(* IEC 61131-3 sources: rusty/tests/lit/ir_tests, 10 files *)

(* ---- adr_ptr_arith.st ---- *)
// RUN: %COMPILE_IR %s | %CHECK_IR %s
//
// Structural pin for the #1749 fix: `ADR(x) + N` must lower to
// `ptrtoint` + `add` (byte-stride integer arithmetic), not panic. ADR is
// declared `: LWORD` so the binary `+` flows through the integer path; the
// codegen entry now routes pointer operands through
// `convert_to_int_value_if_pointer` (matching the existing comparison-op
// path) instead of an unconditional `into_int_value()` that crashed inkwell.

FUNCTION main
VAR
    arr : ARRAY[0..3] OF BYTE;
    pt  : REF_TO BYTE;
END_VAR

pt := ADR(arr) + 2;
pt^ := BYTE#16#FF;
END_FUNCTION

// CHECK: ptrtoint ptr %{{.*}} to i64
// CHECK-NEXT: add i64 %{{.*}}, 2
// CHECK-NEXT: inttoptr i64 %{{.*}} to ptr

(* ---- var_input_aggregate_pass_by_ref.st ---- *)
// RUN: %COMPILE_IR %s | %CHECK_IR %s

// Aggregate VAR_INPUT arguments must be passed by pointer; emitting
// `bitcast ptr -> [N x T]` is invalid IR. See #1718.

FUNCTION foo
   VAR_INPUT
       arr : ARRAY[1..3] OF DINT;
   END_VAR
END_FUNCTION

FUNCTION main
   foo([1, 2, 3]);
END_FUNCTION

// CHECK-LABEL: define {{.*}}@main
// CHECK:       %{{[a-zA-Z0-9_.]+}} = alloca [3 x i32]
// CHECK:       store [3 x i32]
// CHECK:       call {{.*}}@foo(ptr {{.*}})
// CHECK-NOT:   bitcast ptr {{.*}} to [

(* ---- variadic_null_terminator.st ---- *)
// RUN: %COMPILE_IR %s | %CHECK_IR %s
//
// Calls to untyped C-style variadics (`args : ...`) carry an implicit null pointer as their
// last argument. The callee has no way of its own to know how many arguments it received, so
// APIs that walk the list until a terminator read past the arguments without it. Format- and
// count-directed callees read only the arguments they expect and never see the terminator.
//
// Typed variadics keep their argument list unchanged: a `{sized} T...` passes (count, array)
// and a typed unsized `T...` has a concrete callee signature, so a terminator would corrupt
// the contract in both cases.

{external}
FUNCTION untyped : DINT
VAR_INPUT
    fmt : STRING;
    args : ...;
END_VAR
END_FUNCTION

{external}
FUNCTION typed : DINT
VAR_INPUT
    count : DINT;
    args : DINT...;
END_VAR
END_FUNCTION

{external}
FUNCTION sized : DINT
VAR_INPUT
    args : {sized} DINT...;
END_VAR
END_FUNCTION

FUNCTION main : DINT
VAR
    text : STRING := 'text';
END_VAR
    // A call without any variadic argument is still terminated. This is the case in which a
    // terminator-based callee reads past the argument list without the terminator.
    untyped(text);
    // CHECK: call i32 (ptr, ...) @untyped(ptr {{.*}}, ptr null)

    untyped(text, DINT#1, DINT#2);
    // CHECK: call i32 (ptr, ...) @untyped(ptr {{.*}}, i32 1, i32 2, ptr null)

    // The `, !dbg` suffix pins the end of the argument list, so an added terminator fails here.
    typed(DINT#2, DINT#1, DINT#2);
    // CHECK: call i32 (i32, ...) @typed(i32 2, i32 1, i32 2), !dbg

    sized(DINT#1, DINT#2, DINT#3);
    // CHECK: call i32 @sized(i32 3, ptr {{.*}}), !dbg
END_FUNCTION

(* ---- action_call_stores_var_in_out_address.st ---- *)
// RUN: %COMPILE_IR %s | %CHECK_IR %s
//
// Pin the IR shape that the #1576 fix (commit 2b3388f) put in place: when
// calling an action that inherits a `VAR_IN_OUT` from its parent FB, the
// caller must (a) GEP to the FB's in-out slot and (b) store the local's
// address there before invoking the action. Skipping either step leaves the
// pointer NULL and the action segfaults at runtime — runtime coverage lives
// in `tests/lit/single/actions/action_call_with_var_in_out.st`; this test
// is the structural guardrail.

PROGRAM mainProg
VAR
    fb : fb_t;
    localBool : BOOL;
END_VAR
    fb.foo(myInOut := localBool);
END_PROGRAM

FUNCTION_BLOCK fb_t
VAR_IN_OUT
    myInOut : BOOL;
END_VAR
END_FUNCTION_BLOCK

ACTIONS
    ACTION foo
        myInOut := myInOut;
    END_ACTION
END_ACTIONS

// CHECK-LABEL: define void @mainProg(
// CHECK: %fb = getelementptr inbounds nuw %mainProg, {{.*}}, i32 0, i32 0
// CHECK: %localBool = getelementptr inbounds nuw %mainProg, {{.*}}, i32 0, i32 1
// CHECK: getelementptr inbounds %fb_t, ptr %fb, i32 0, i32 1
// CHECK-NEXT: store ptr %localBool, ptr {{%[0-9]+}}, align 8
// CHECK-NEXT: call void @fb_t__foo(ptr %fb)

(* ---- external_fb_array_const_init.st ---- *)
// RUN: %COMPILE_IR --generate-external-constructors %s | %CHECK_IR %s
//
// When an {external} function block has an array with a constant initializer,
// compiling with --generate-external-constructors should:
//   1. Produce a .const_init global for the array
//   2. Define (not declare) the ctor
//   3. Use memcpy from the .const_init in the ctor body

{external}
FUNCTION_BLOCK myFb
VAR
    arr : ARRAY[0..4] OF DINT := [1, 2, 3, 4, 5];
END_VAR
END_FUNCTION_BLOCK

PROGRAM Main
VAR
    fb : myFb;
END_VAR
END_PROGRAM

// The const_init global should exist for the array
// CHECK: @.const_init = private unnamed_addr constant [5 x i32] [i32 1, i32 2, i32 3, i32 4, i32 5]

// The ctor for myFb should be defined (has body), not just declared
// CHECK: define void @myFb__ctor(ptr %0)

// The ctor should use memcpy from the const_init
// CHECK: call void @llvm.memcpy{{.*}}@.const_init

(* ---- external_fb_array_no_init_globals.st ---- *)
// RUN: %COMPILE_IR %s | %CHECK_IR %s
//
// When an {external} function block has an array with a constant initializer,
// compiling WITHOUT --generate-external-constructors should:
//   1. NOT produce any .const_init or __init globals for the external FB
//   2. Declare (not define) the ctor

{external}
FUNCTION_BLOCK myFb
VAR
    arr : ARRAY[0..4] OF DINT := [1, 2, 3, 4, 5];
END_VAR
END_FUNCTION_BLOCK

PROGRAM Main
VAR
    fb : myFb;
END_VAR
END_PROGRAM

// No .const_init or __myFb.arr__init globals should be present.
// CHECK-NOT directives must come before CHECK to scan from start of input.
// CHECK-NOT: @.const_init
// CHECK-NOT: @__myFb.arr__init

// The ctor for myFb should be declared (external), not defined
// CHECK: declare void @myFb__ctor(ptr)

(* ---- fb_call_no_int_extension_attrs.st ---- *)
// REQUIRES: host-x86_64
// RUN: %COMPILE_IR %s | %CHECK_IR %s
//
// Direct FUNCTION_BLOCK invocations (e.g. `myFbInstance(in_val := …)`) lower to
// a gep+store of each argument into the instance struct followed by a call to
// the FB body that takes only the instance pointer — there are no scalar
// arguments in the LLVM call signature, so no `signext`/`zeroext` attribute is
// applicable. Regression for #1146 review feedback: confirms the call-side
// integer-extension pass leaves direct FB calls alone.
//
// Gated to host-x86_64 to mirror sub32_int_ffi_extension.st: `signext`/`zeroext`
// are only emitted on x86 family and Apple/Darwin targets. The point of this
// test is the *absence* of those tokens, but on AAPCS targets they would be
// absent for a different reason (target gate), which would make the test
// trivially green and hide a future regression on x86.

FUNCTION_BLOCK myFb
VAR_INPUT
    in_val : SINT;
END_VAR
END_FUNCTION_BLOCK

PROGRAM main
VAR
    instance : myFb;
END_VAR
    instance(in_val := SINT#-1);
END_PROGRAM

// The body call passes only the instance struct pointer (LLVM 21 opaque
// `ptr`) — no `signext`/`zeroext` token should appear on the call line.
// CHECK: call void @myFb(ptr {{.*}})
// CHECK-NOT: call void @myFb({{.*}}signext{{.*}})
// CHECK-NOT: call void @myFb({{.*}}zeroext{{.*}})

(* ---- included_struct_ctor.st ---- *)
// RUN: %COMPILE_IR -i %p/include/included_types.st %s | %CHECK_IR %s

PROGRAM Main
VAR
    s : IncludedStruct;
END_VAR
END_PROGRAM

// The declaration may precede or follow Main__ctor depending on the unit order
// CHECK-NOT: define{{.*}}@IncludedStruct__ctor
// CHECK-DAG: define void @Main__ctor(ptr %0) {
// CHECK-DAG: call void @IncludedStruct__ctor(ptr %s)
// CHECK-DAG: declare void @IncludedStruct__ctor(ptr)
// CHECK-NOT: define{{.*}}@IncludedStruct__ctor

(* ---- nested_array_const_expression_init.st ---- *)
// RUN: %COMPILE_IR %s | %CHECK_IR %s
//
// Structural pin for the PRG-4521 fix: constant expressions inside nested
// array initializers are const-folded, so the initializer lowers to a folded
// constant global copied via memcpy. Previously the raw expression tree
// reached codegen's literal generator and failed with "Cannot generate
// Literal for BinaryExpression". Runtime coverage lives in
// tests/lit/single/init/array_const_expression_init.st.

PROGRAM mainProg
VAR
    mArr : ARRAY[0..1] OF ARRAY[0..1] OF UDINT := [[UDINT#0 + UDINT#1, UDINT#0], [UDINT#0, UDINT#2 - UDINT#1]];
END_VAR
    ;
END_PROGRAM

// The type's __init global is fully folded to [1, 0], [0, 1].
// CHECK: @__mainProg.mArr__init = unnamed_addr constant [2 x [2 x i32]] {{\[}}[2 x i32] [i32 1, i32 0], [2 x i32] [i32 0, i32 1]]

// The ctor assignment is folded as well and copied via memcpy.
// CHECK: @.const_init = private unnamed_addr constant [2 x [2 x i32]] {{\[}}[2 x i32] [i32 1, i32 0], [2 x i32] [i32 0, i32 1]]
// CHECK: define void @mainProg__ctor(ptr %0)
// CHECK: call void @llvm.memcpy{{.*}}@.const_init

(* ---- sub32_int_ffi_extension.st ---- *)
// REQUIRES: host-x86_64
// RUN: %COMPILE_IR %s | %CHECK_IR %s
//
// Regression for #1146. Verify call sites and declarations of functions taking sub-32-bit
// integer parameters carry the correct LLVM `signext`/`zeroext` parameter attributes.
// Without these, optimized release builds of FFI'd callees (e.g. the Rust stdlib) read
// garbage upper register bits instead of the intended signed value — see also
// `cargo test --release -p iec61131std mul_ltime_signed`.
//
// Gated to host-x86_64 because the codegen emission is target-aware: x86 family and
// Apple/Darwin emit the attributes; plain AAPCS (aarch64-unknown-linux-gnu) does not
// and the FILECHECK lines below would not match. The runtime regression coverage for
// the AAPCS path lives under tests/lit/single/stdlib_overflow/sub32_ffi_return_*.st.

{external}
FUNCTION extFunc : LINT
VAR_INPUT
    in1 : SINT;
    in2 : USINT;
    in3 : INT;
    in4 : UINT;
    in5 : BOOL;
END_VAR
END_FUNCTION

PROGRAM main
VAR
    a : LINT;
END_VAR
    a := extFunc(SINT#-1, USINT#1, INT#-1, UINT#1, FALSE);
END_PROGRAM

// BOOL is lowered to `i8` at the FFI boundary, not `i1`; both still get `zeroext`.
// `CHECK-DAG` so the order of `call`/`declare` (call first under --debug, declare last)
// doesn't matter to this test.
// CHECK-DAG: call i64 @extFunc(i8 signext {{.*}}, i8 zeroext {{.*}}, i16 signext {{.*}}, i16 zeroext {{.*}}, i8 zeroext {{.*}})
// CHECK-DAG: declare i64 @extFunc(i8 signext, i8 zeroext, i16 signext, i16 zeroext, i8 zeroext)
